PROGRAM prg_Safety
VAR
	(*
	rt_TSafe_OK: R_TRIG;
	rt_TSafe_Err: R_TRIG;
	ton_TSafe_OK: TON;
	ton_TSafe_Err_Reset_ON: TON;
	ton_TSafe_Err_Reset_OFF: TON;
	*)
	fbTwinSAFE: ARRAY[1..1] OF FB_TwinSAFE;
	
	HMI_ES1_Restart: BOOL;
	HMI_ES2_Restart: BOOL;
	HMI_ES3_Restart: BOOL;
	HMI_ES4_Restart: BOOL;
	
	rtStateSafe: R_TRIG;
	ftStateSafe: F_TRIG;
END_VAR


act_Call_TSs();


{IF defined (Production)}
	bStateSafe_ES1:=arSafe[1].stSafetyIn.ES1_State;
	//bStateSafe_ES2:=arSafe[1].stSafetyIn.ES2_State;
	bStateSafe_ES3:=arSafe[1].stSafetyIn.ES3_State;
	//bStateSafe_ES4:=arSafe[1].stSafetyIn.ES4_State;
{ELSIF defined (Simulation_IO)}
	bES_Bypass:= TRUE;

	bStateSafe_ES1:=TRUE;
	bStateSafe_ES2:=TRUE;
	bStateSafe_ES3:=TRUE;
	bStateSafe_ES4:=TRUE;
{END_IF}

IF TRUE 
AND bStateSafe_ES1
//AND bStateSafe_ES2
AND bStateSafe_ES3
//AND bStateSafe_ES4

OR bES_Bypass

THEN;
	bStateSafe:=TRUE;
ELSE;
	bStateSafe:=FALSE;
END_IF
rtStateSafe(CLK:=bStateSafe);
ftStateSafe(CLK:=bStateSafe);

IF bStateSafe THEN
	sBitmap_ESButton:= 'ImagePool.EStop_OK2';
	stBitMap:='bitmap\EStop_OK2.bmp';
ELSE
	sBitmap_ESButton:= 'ImagePool.EStop_ACT2';
	stBitMap:='bitmap\EStop_ACT2.bmp';
END_IF

(*
ton_TSafe_OK(IN:=g_IO.TSafeIn.InRun AND NOT g_IO.TSafeIn.COM_Err, PT:=T#1S );
IF ton_TSafe_OK.Q THEN;
	bStateSafe:=TRUE;
ELSE;
	bStateSafe:=FALSE;	
END_IF
rt_TSafe_OK(CLK:=ton_TSafe_OK.Q );
IF rt_TSafe_OK.Q THEN;
	m_Print_Success_Message();
END_IF



rt_TSafe_Err(CLK:=g_IO.TSafeIn.COM_Err);
IF rt_TSafe_Err.Q THEN;
	m_Print_Error_Message();
END_IF

ton_TSafe_Err_Reset_ON(IN:=g_IO.TSafeIn.COM_Err AND NOT g_IO.TSafeOut.ErrACK, PT:=T#2S );
IF ton_TSafe_Err_Reset_ON.Q THEN;
	g_IO.TSafeOut.ErrACK:=TRUE;
END_IF

ton_TSafe_Err_Reset_OFF(IN:=g_IO.TSafeOut.ErrACK, PT:=T#1S );
IF ton_TSafe_Err_Reset_OFF.Q THEN;
	g_IO.TSafeOut.ErrACK:=FALSE;
END_IF
*)

ACTION act_Call_TSs:
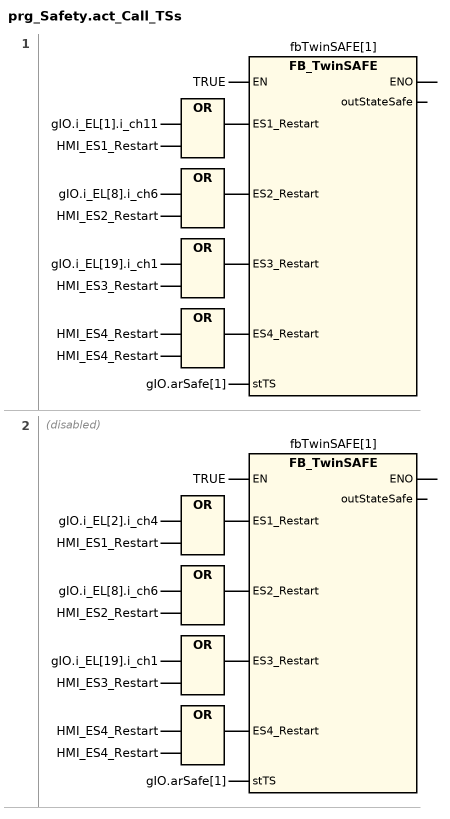
// NETWORK 1
fbTwinSAFE[1](
    ES1_Restart := gIO.i_EL[1].i_ch11 OR HMI_ES1_Restart,
    ES2_Restart := gIO.i_EL[8].i_ch6 OR HMI_ES2_Restart,
    ES3_Restart := gIO.i_EL[19].i_ch1 OR HMI_ES3_Restart,
    ES4_Restart := HMI_ES4_Restart OR HMI_ES4_Restart,
    stTS := gIO.arSafe[1]); // FB_TwinSAFE

// NETWORK 2 (disabled)
// fbTwinSAFE[1](
//     ES1_Restart := gIO.i_EL[2].i_ch4 OR HMI_ES1_Restart,
//     ES2_Restart := gIO.i_EL[8].i_ch6 OR HMI_ES2_Restart,
//     ES3_Restart := gIO.i_EL[19].i_ch1 OR HMI_ES3_Restart,
//     ES4_Restart := HMI_ES4_Restart OR HMI_ES4_Restart,
//     stTS := gIO.arSafe[1]); // FB_TwinSAFE
END_ACTION

METHOD m_Print_Error_Message : BOOL
VAR_INPUT
END_VAR

VAR
	i: INT;
	sActErrorID: STRING(11);
	sModuleDescription: STRING(80);
END_VAR

sActErrorID:='0x999x0';
sModuleDescription:='TwinSAFE Group';

FOR i:=100 TO 2 BY -1 DO
	Buffer_Act_Message[i]:=Buffer_Act_Message[i-1];
END_FOR

Buffer_Act_Message[1].sDateTime:=sRealTime_Date;
Buffer_Act_Message[1].sErrID:=sActErrorID;
Buffer_Act_Message[1].sModuleDescription:=sModuleDescription;
Buffer_Act_Message[1].sLevel:='Error';
Buffer_Act_Message[1].sErrorMessage:='';

Buffer_Act_Message[1].sErrorMessage:=CONCAT(Buffer_Act_Message[1].sErrorMessage,'TwinSAFE group has a communication error');
FUN_Write_Line_To_History();
END_METHOD

METHOD m_Print_Success_Message : BOOL
VAR_INPUT
END_VAR

VAR
	i: INT;
	sActErrorID: STRING(11);
	sModuleDescription: STRING(80);
END_VAR

sActErrorID:='0x999x0';
sModuleDescription:='TwinSAFE Group';

FOR i:=1000 TO 2 BY -1 DO
	Buffer_Act_History[i]:=Buffer_Act_History[i-1];
END_FOR

Buffer_Act_History[1].sDateTime:=sRealTime_Date;
Buffer_Act_History[1].sErrID:=sActErrorID;
Buffer_Act_History[1].sModuleDescription:=sModuleDescription;
Buffer_Act_History[1].sLevel:='Message';
Buffer_Act_History[1].sErrorMessage:='';

Buffer_Act_History[1].sErrorMessage:=CONCAT(Buffer_Act_History[1].sErrorMessage,'TwinSAFE state is OK');
END_METHOD

END_PROGRAM

(* stored: Version 1.1.0.1, ProductVersion 3.1.4026.21
   POU prg_Safety: Id {db89eb8b-da04-4986-84d3-a7f6079fbab6}, SpecialFunc None
   Action act_Call_TSs: Id {bb85fd28-de4b-415c-82fd-1939945fdd5f}
   Method m_Print_Error_Message: Id {6a416efc-1748-4d8e-9420-3cb4c1f658da}
   Method m_Print_Success_Message: Id {ea77dc15-18d3-4625-bca6-cfe5f939b2cc} *)
